(* Logix 5000 project; controller CIP vendor 1 type 14 code 106 rev 20.12; software revision 20.06; part 4 of 13 *)
(* tags used below, declared in another part *)
   Alarm_Ack : INT[8];
   Alarm_Present : INT[8];
   Alarm_Remote_Ack_All : BOOL;
   Alarm_Timer : TIMER[128];
   Bit : BOOL[128];
   IO_Status : INT;
   IO_Status_Masked : INT;
   Level_Bits : BOOL[32];
   Level_Timers : TIMER[20];
   OpCode_Pin : DINT[5];
   Recipe : RECIPE[41];
   SCLD_Dryer_Duct_Temp : REAL;
   SCLD_Solution_Tank_Lvl : REAL;
   SCLD_Supply_Flow : REAL;
   SCLD_Supply_Flow_CIP100 : REAL;
   SCLD_Supply_Flow_CIP200 : REAL;
   SCLD_Supply_Pressure : REAL;
   SCLD_Supply_Temp : REAL;
   Timer : TIMER[99];
   Timer_Chem1_Pump : TIMER[7];
   Timer_Chem2_Pump : TIMER[7];
(* MainProgram, continued *)

ROUTINE _05_ALARMS   (* ladder *)
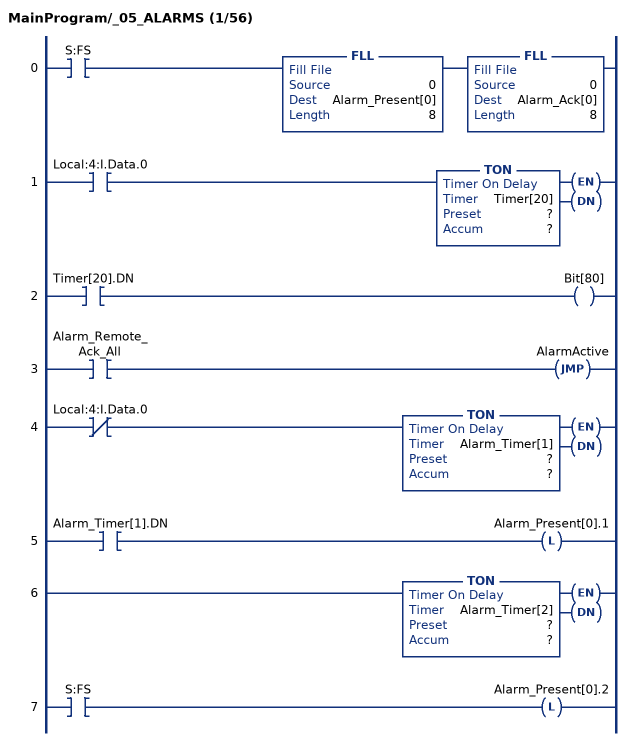
   0: XIC(S:FS)FLL(0,Alarm_Present[0],8)FLL(0,Alarm_Ack[0],8);
   1: XIC(Local:4:I.Data.0)TON(Timer[20],?,?);
   2: XIC(Timer[20].DN)OTE(Bit[80]);
   3: XIC(Alarm_Remote_Ack_All)JMP(AlarmActive);
   4: XIO(Local:4:I.Data.0)TON(Alarm_Timer[1],?,?);
   5: XIC(Alarm_Timer[1].DN)OTL(Alarm_Present[0].1);
   6: TON(Alarm_Timer[2],?,?);
   7: XIC(S:FS)OTL(Alarm_Present[0].2);
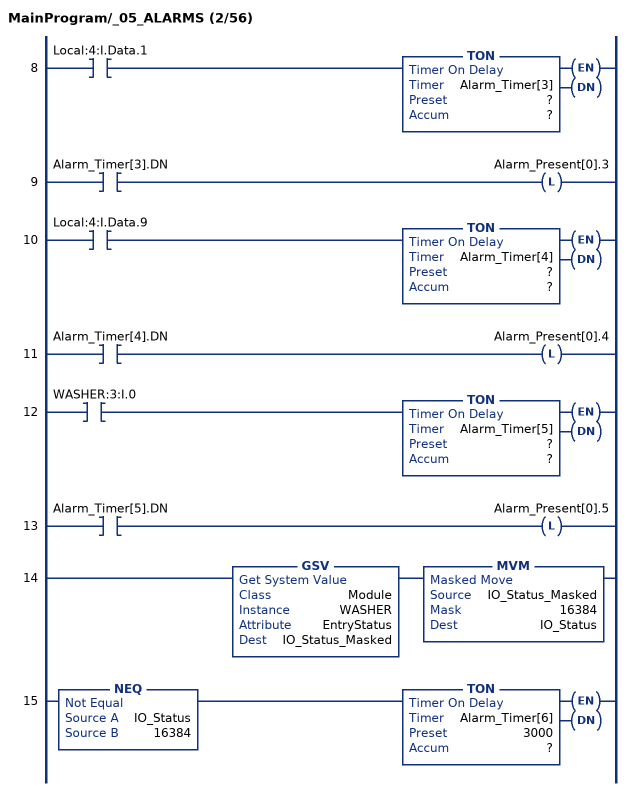
   8: XIC(Local:4:I.Data.1)TON(Alarm_Timer[3],?,?);
   9: XIC(Alarm_Timer[3].DN)OTL(Alarm_Present[0].3);
   10: XIC(Local:4:I.Data.9)TON(Alarm_Timer[4],?,?);
   11: XIC(Alarm_Timer[4].DN)OTL(Alarm_Present[0].4);
   12: XIC(WASHER:3:I.0)TON(Alarm_Timer[5],?,?);
   13: XIC(Alarm_Timer[5].DN)OTL(Alarm_Present[0].5);
   14: GSV(Module,WASHER,EntryStatus,IO_Status_Masked)MVM(IO_Status_Masked,16384,IO_Status);
   15: NEQ(IO_Status,16384)TON(Alarm_Timer[6],?,?);
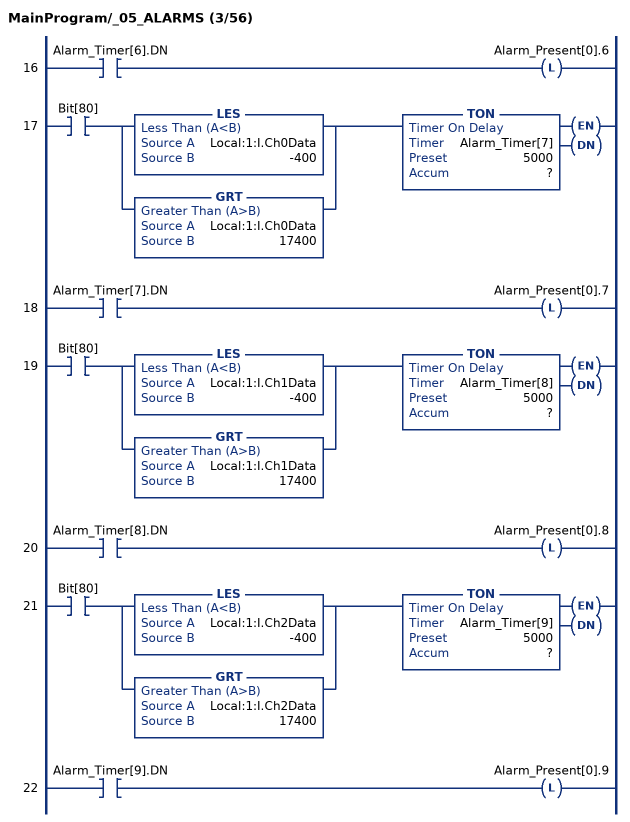
   16: XIC(Alarm_Timer[6].DN)OTL(Alarm_Present[0].6);
   17: XIC(Bit[80])[LES(Local:1:I.Ch0Data,-400) ,GRT(Local:1:I.Ch0Data,17400) ]TON(Alarm_Timer[7],?,?);
   18: XIC(Alarm_Timer[7].DN)OTL(Alarm_Present[0].7);
   19: XIC(Bit[80])[LES(Local:1:I.Ch1Data,-400) ,GRT(Local:1:I.Ch1Data,17400) ]TON(Alarm_Timer[8],?,?);
   20: XIC(Alarm_Timer[8].DN)OTL(Alarm_Present[0].8);
   21: XIC(Bit[80])[LES(Local:1:I.Ch2Data,-400) ,GRT(Local:1:I.Ch2Data,17400) ]TON(Alarm_Timer[9],?,?);
   22: XIC(Alarm_Timer[9].DN)OTL(Alarm_Present[0].9);
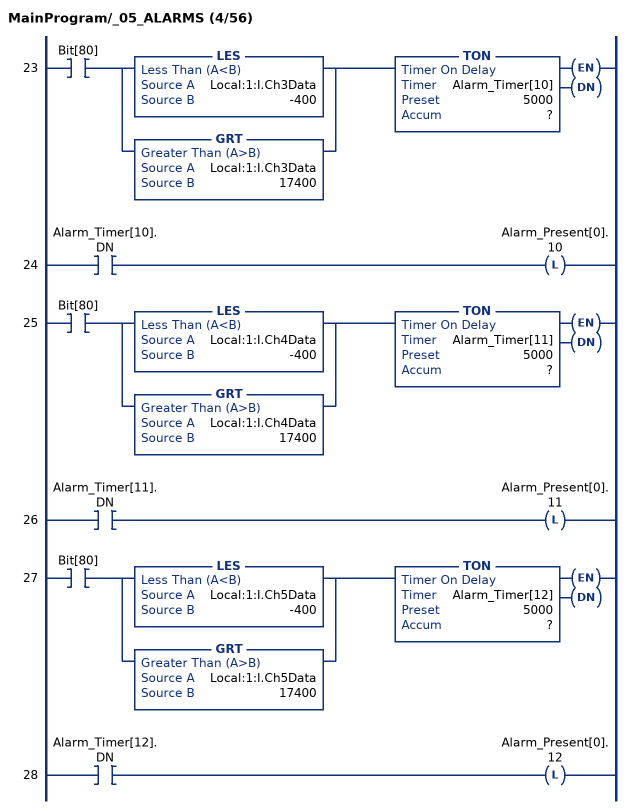
   23: XIC(Bit[80])[LES(Local:1:I.Ch3Data,-400) ,GRT(Local:1:I.Ch3Data,17400) ]TON(Alarm_Timer[10],?,?);
   24: XIC(Alarm_Timer[10].DN)OTL(Alarm_Present[0].10);
   25: XIC(Bit[80])[LES(Local:1:I.Ch4Data,-400) ,GRT(Local:1:I.Ch4Data,17400) ]TON(Alarm_Timer[11],?,?);
   26: XIC(Alarm_Timer[11].DN)OTL(Alarm_Present[0].11);
   27: XIC(Bit[80])[LES(Local:1:I.Ch5Data,-400) ,GRT(Local:1:I.Ch5Data,17400) ]TON(Alarm_Timer[12],?,?);
   28: XIC(Alarm_Timer[12].DN)OTL(Alarm_Present[0].12);
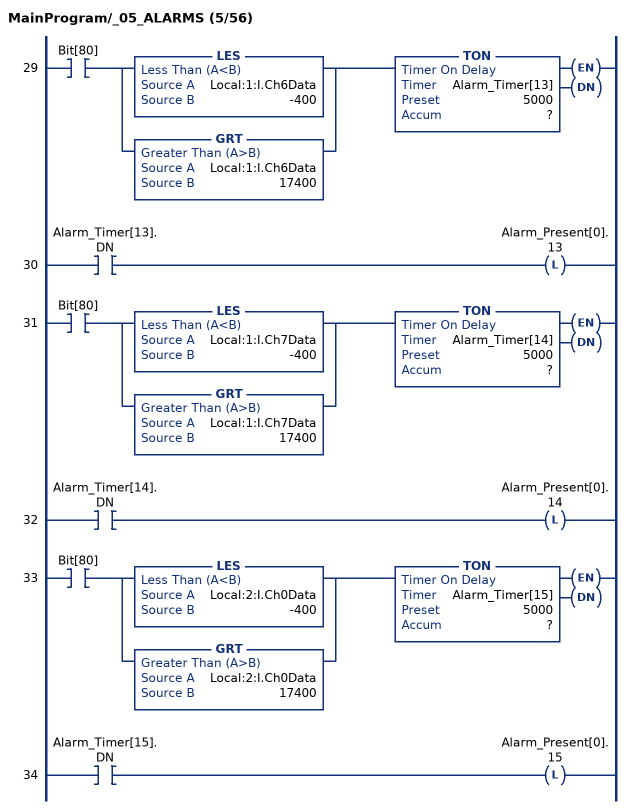
   29: XIC(Bit[80])[LES(Local:1:I.Ch6Data,-400) ,GRT(Local:1:I.Ch6Data,17400) ]TON(Alarm_Timer[13],?,?);
   30: XIC(Alarm_Timer[13].DN)OTL(Alarm_Present[0].13);
   31: XIC(Bit[80])[LES(Local:1:I.Ch7Data,-400) ,GRT(Local:1:I.Ch7Data,17400) ]TON(Alarm_Timer[14],?,?);
   32: XIC(Alarm_Timer[14].DN)OTL(Alarm_Present[0].14);
   33: XIC(Bit[80])[LES(Local:2:I.Ch0Data,-400) ,GRT(Local:2:I.Ch0Data,17400) ]TON(Alarm_Timer[15],?,?);
   34: XIC(Alarm_Timer[15].DN)OTL(Alarm_Present[0].15);
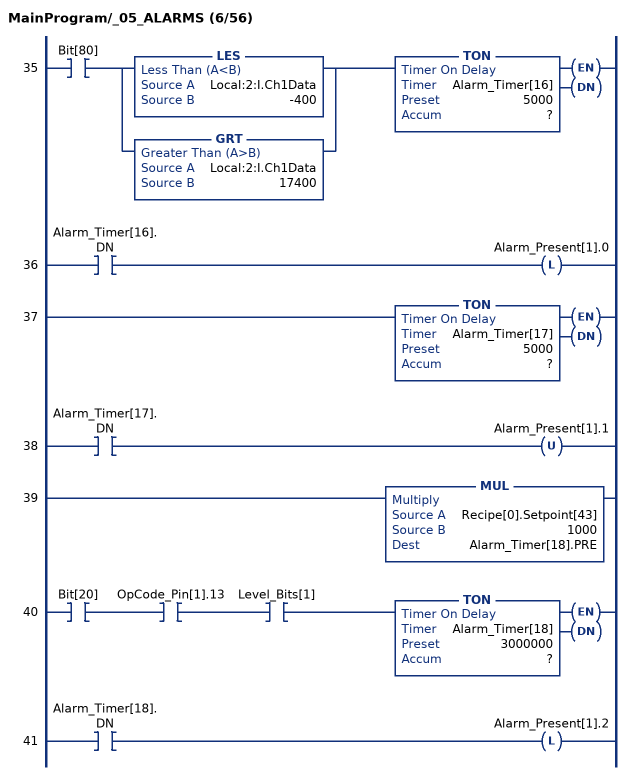
   35: XIC(Bit[80])[LES(Local:2:I.Ch1Data,-400) ,GRT(Local:2:I.Ch1Data,17400) ]TON(Alarm_Timer[16],?,?);
   36: XIC(Alarm_Timer[16].DN)OTL(Alarm_Present[1].0);
   37: TON(Alarm_Timer[17],?,?);
   38: XIC(Alarm_Timer[17].DN)OTU(Alarm_Present[1].1);
   39: MUL(Recipe[0].Setpoint[43],1000,Alarm_Timer[18].PRE);
   40: XIC(Bit[20])XIC(OpCode_Pin[1].13)XIC(Level_Bits[1])TON(Alarm_Timer[18],?,?);
   41: XIC(Alarm_Timer[18].DN)OTL(Alarm_Present[1].2);
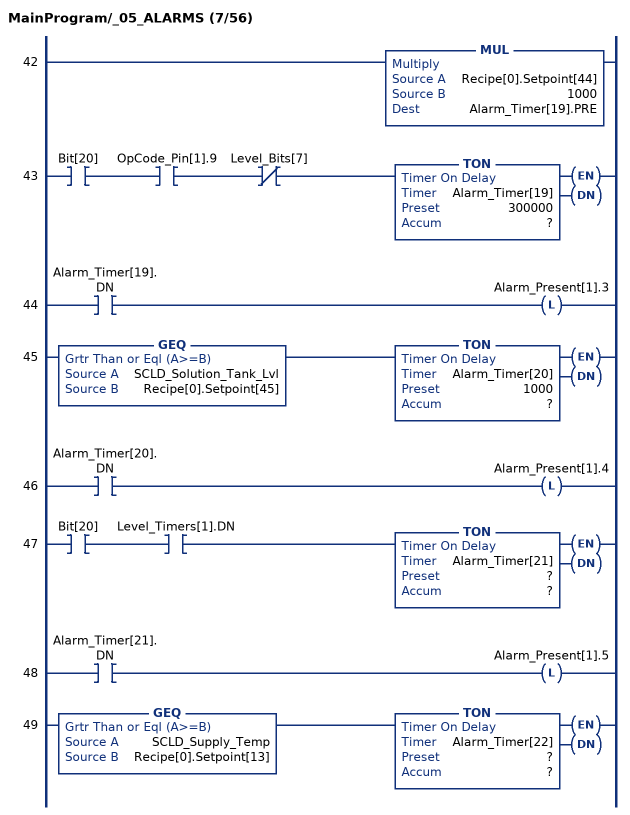
   42: MUL(Recipe[0].Setpoint[44],1000,Alarm_Timer[19].PRE);
   43: XIC(Bit[20])XIC(OpCode_Pin[1].9)XIO(Level_Bits[7])TON(Alarm_Timer[19],?,?);
   44: XIC(Alarm_Timer[19].DN)OTL(Alarm_Present[1].3);
   45: GEQ(SCLD_Solution_Tank_Lvl,Recipe[0].Setpoint[45])TON(Alarm_Timer[20],?,?);
   46: XIC(Alarm_Timer[20].DN)OTL(Alarm_Present[1].4);
   47: XIC(Bit[20])XIC(Level_Timers[1].DN)TON(Alarm_Timer[21],?,?);
   48: XIC(Alarm_Timer[21].DN)OTL(Alarm_Present[1].5);
   49: GEQ(SCLD_Supply_Temp,Recipe[0].Setpoint[13])TON(Alarm_Timer[22],?,?);
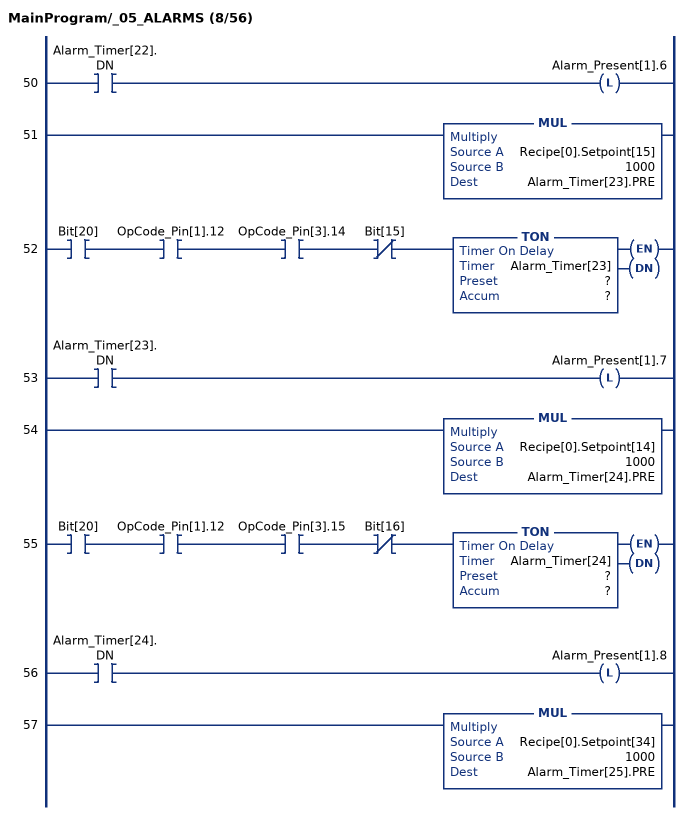
   50: XIC(Alarm_Timer[22].DN)OTL(Alarm_Present[1].6);
   51: MUL(Recipe[0].Setpoint[15],1000,Alarm_Timer[23].PRE);
   52: XIC(Bit[20])XIC(OpCode_Pin[1].12)XIC(OpCode_Pin[3].14)XIO(Bit[15])TON(Alarm_Timer[23],?,?);
   53: XIC(Alarm_Timer[23].DN)OTL(Alarm_Present[1].7);
   54: MUL(Recipe[0].Setpoint[14],1000,Alarm_Timer[24].PRE);
   55: XIC(Bit[20])XIC(OpCode_Pin[1].12)XIC(OpCode_Pin[3].15)XIO(Bit[16])TON(Alarm_Timer[24],?,?);
   56: XIC(Alarm_Timer[24].DN)OTL(Alarm_Present[1].8);
   57: MUL(Recipe[0].Setpoint[34],1000,Alarm_Timer[25].PRE);
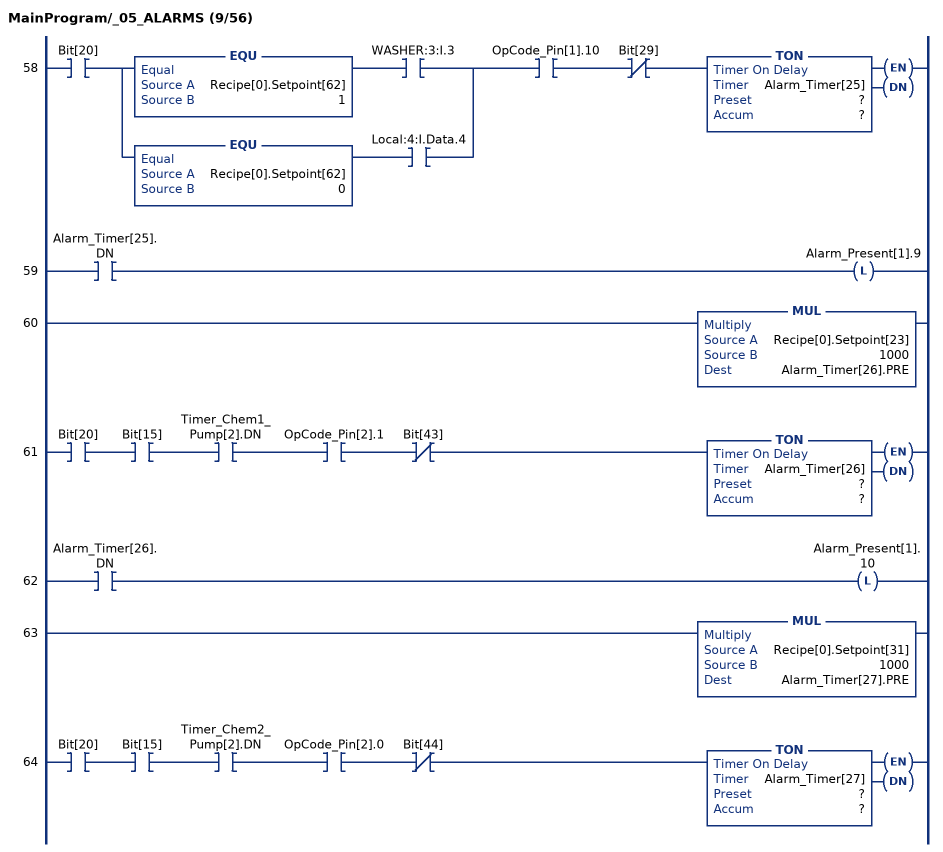
   58: XIC(Bit[20])[EQU(Recipe[0].Setpoint[62],1) XIC(WASHER:3:I.3) ,EQU(Recipe[0].Setpoint[62],0) XIC(Local:4:I.Data.4) ]XIC(OpCode_Pin[1].10)XIO(Bit[29])TON(Alarm_Timer[25],?,?);
   59: XIC(Alarm_Timer[25].DN)OTL(Alarm_Present[1].9);
   60: MUL(Recipe[0].Setpoint[23],1000,Alarm_Timer[26].PRE);
   61: XIC(Bit[20])XIC(Bit[15])XIC(Timer_Chem1_Pump[2].DN)XIC(OpCode_Pin[2].1)XIO(Bit[43])TON(Alarm_Timer[26],?,?);
   62: XIC(Alarm_Timer[26].DN)OTL(Alarm_Present[1].10);
   63: MUL(Recipe[0].Setpoint[31],1000,Alarm_Timer[27].PRE);
   64: XIC(Bit[20])XIC(Bit[15])XIC(Timer_Chem2_Pump[2].DN)XIC(OpCode_Pin[2].0)XIO(Bit[44])TON(Alarm_Timer[27],?,?);
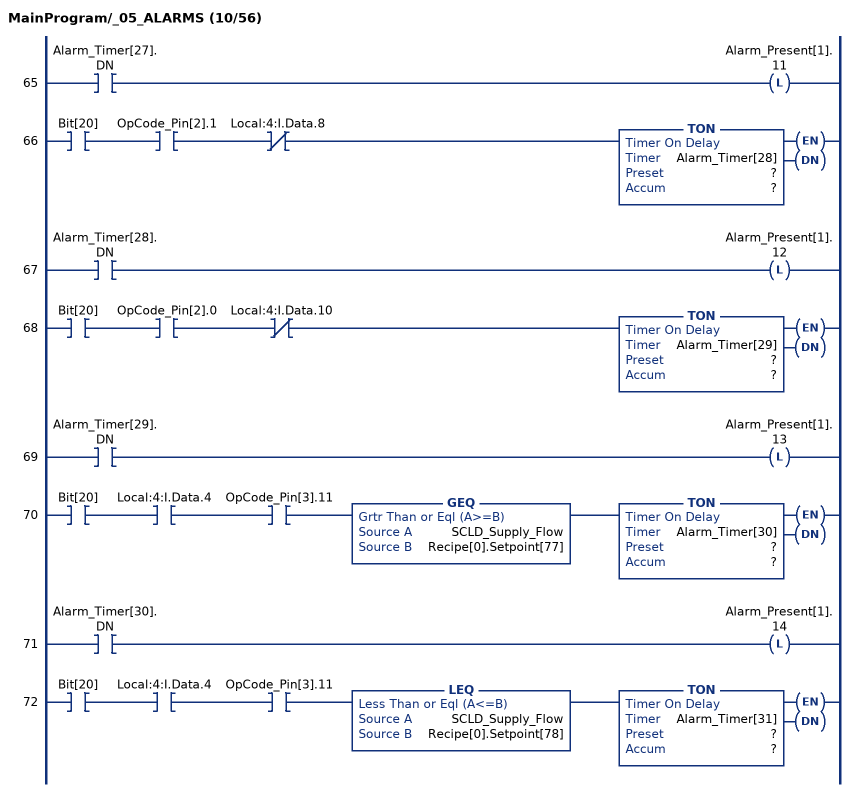
   65: XIC(Alarm_Timer[27].DN)OTL(Alarm_Present[1].11);
   66: XIC(Bit[20])XIC(OpCode_Pin[2].1)XIO(Local:4:I.Data.8)TON(Alarm_Timer[28],?,?);
   67: XIC(Alarm_Timer[28].DN)OTL(Alarm_Present[1].12);
   68: XIC(Bit[20])XIC(OpCode_Pin[2].0)XIO(Local:4:I.Data.10)TON(Alarm_Timer[29],?,?);
   69: XIC(Alarm_Timer[29].DN)OTL(Alarm_Present[1].13);
   70: XIC(Bit[20])XIC(Local:4:I.Data.4)XIC(OpCode_Pin[3].11)GEQ(SCLD_Supply_Flow,Recipe[0].Setpoint[77])TON(Alarm_Timer[30],?,?);
   71: XIC(Alarm_Timer[30].DN)OTL(Alarm_Present[1].14);
   72: XIC(Bit[20])XIC(Local:4:I.Data.4)XIC(OpCode_Pin[3].11)LEQ(SCLD_Supply_Flow,Recipe[0].Setpoint[78])TON(Alarm_Timer[31],?,?);
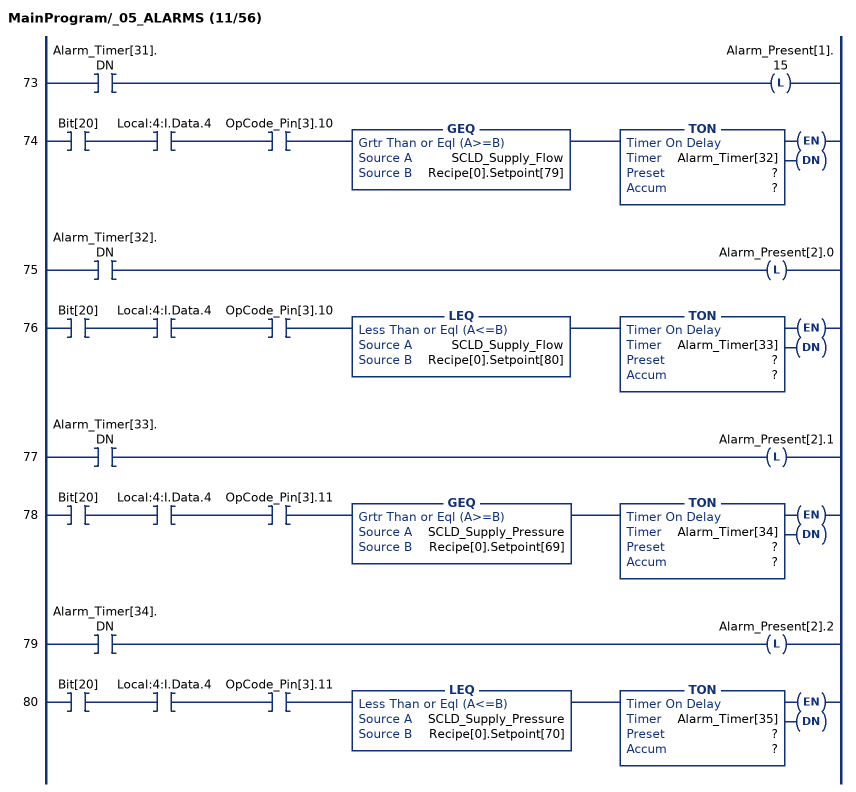
   73: XIC(Alarm_Timer[31].DN)OTL(Alarm_Present[1].15);
   74: XIC(Bit[20])XIC(Local:4:I.Data.4)XIC(OpCode_Pin[3].10)GEQ(SCLD_Supply_Flow,Recipe[0].Setpoint[79])TON(Alarm_Timer[32],?,?);
   75: XIC(Alarm_Timer[32].DN)OTL(Alarm_Present[2].0);
   76: XIC(Bit[20])XIC(Local:4:I.Data.4)XIC(OpCode_Pin[3].10)LEQ(SCLD_Supply_Flow,Recipe[0].Setpoint[80])TON(Alarm_Timer[33],?,?);
   77: XIC(Alarm_Timer[33].DN)OTL(Alarm_Present[2].1);
   78: XIC(Bit[20])XIC(Local:4:I.Data.4)XIC(OpCode_Pin[3].11)GEQ(SCLD_Supply_Pressure,Recipe[0].Setpoint[69])TON(Alarm_Timer[34],?,?);
   79: XIC(Alarm_Timer[34].DN)OTL(Alarm_Present[2].2);
   80: XIC(Bit[20])XIC(Local:4:I.Data.4)XIC(OpCode_Pin[3].11)LEQ(SCLD_Supply_Pressure,Recipe[0].Setpoint[70])TON(Alarm_Timer[35],?,?);
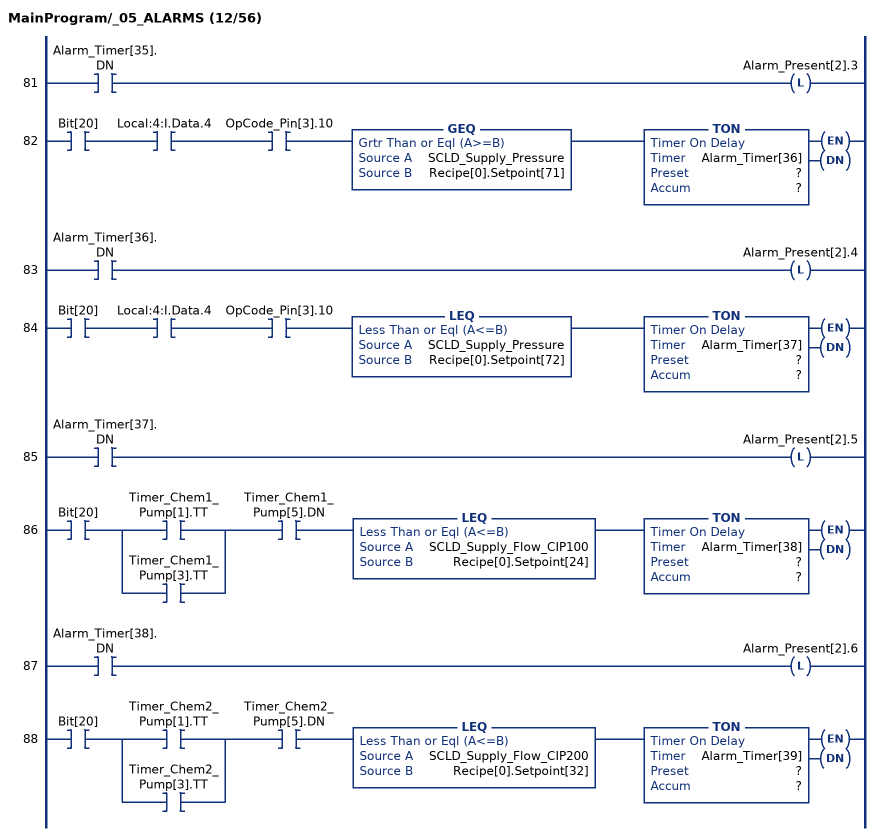
   81: XIC(Alarm_Timer[35].DN)OTL(Alarm_Present[2].3);
   82: XIC(Bit[20])XIC(Local:4:I.Data.4)XIC(OpCode_Pin[3].10)GEQ(SCLD_Supply_Pressure,Recipe[0].Setpoint[71])TON(Alarm_Timer[36],?,?);
   83: XIC(Alarm_Timer[36].DN)OTL(Alarm_Present[2].4);
   84: XIC(Bit[20])XIC(Local:4:I.Data.4)XIC(OpCode_Pin[3].10)LEQ(SCLD_Supply_Pressure,Recipe[0].Setpoint[72])TON(Alarm_Timer[37],?,?);
   85: XIC(Alarm_Timer[37].DN)OTL(Alarm_Present[2].5);
   86: XIC(Bit[20])[XIC(Timer_Chem1_Pump[1].TT) ,XIC(Timer_Chem1_Pump[3].TT) ]XIC(Timer_Chem1_Pump[5].DN)LEQ(SCLD_Supply_Flow_CIP100,Recipe[0].Setpoint[24])TON(Alarm_Timer[38],?,?);
   87: XIC(Alarm_Timer[38].DN)OTL(Alarm_Present[2].6);
   88: XIC(Bit[20])[XIC(Timer_Chem2_Pump[1].TT) ,XIC(Timer_Chem2_Pump[3].TT) ]XIC(Timer_Chem2_Pump[5].DN)LEQ(SCLD_Supply_Flow_CIP200,Recipe[0].Setpoint[32])TON(Alarm_Timer[39],?,?);
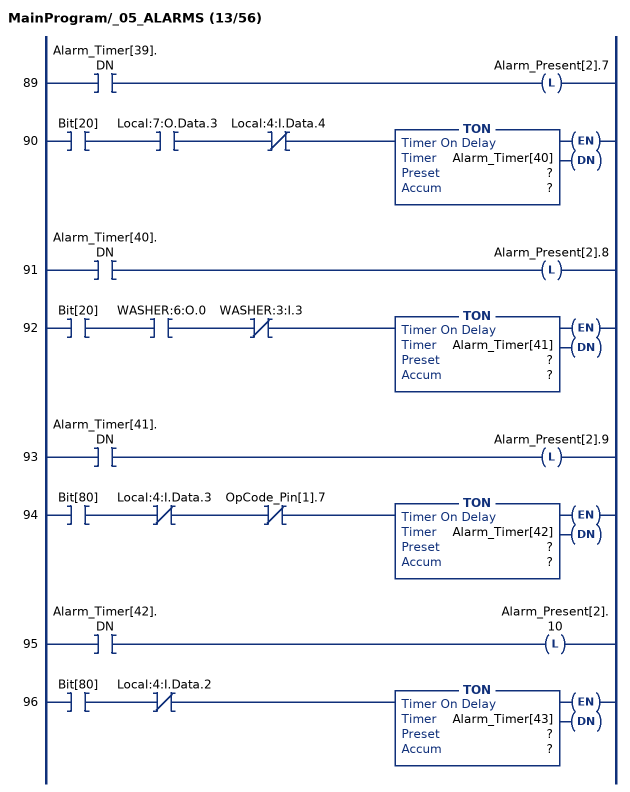
   89: XIC(Alarm_Timer[39].DN)OTL(Alarm_Present[2].7);
   90: XIC(Bit[20])XIC(Local:7:O.Data.3)XIO(Local:4:I.Data.4)TON(Alarm_Timer[40],?,?);
   91: XIC(Alarm_Timer[40].DN)OTL(Alarm_Present[2].8);
   92: XIC(Bit[20])XIC(WASHER:6:O.0)XIO(WASHER:3:I.3)TON(Alarm_Timer[41],?,?);
   93: XIC(Alarm_Timer[41].DN)OTL(Alarm_Present[2].9);
   94: XIC(Bit[80])XIO(Local:4:I.Data.3)XIO(OpCode_Pin[1].7)TON(Alarm_Timer[42],?,?);
   95: XIC(Alarm_Timer[42].DN)OTL(Alarm_Present[2].10);
   96: XIC(Bit[80])XIO(Local:4:I.Data.2)TON(Alarm_Timer[43],?,?);
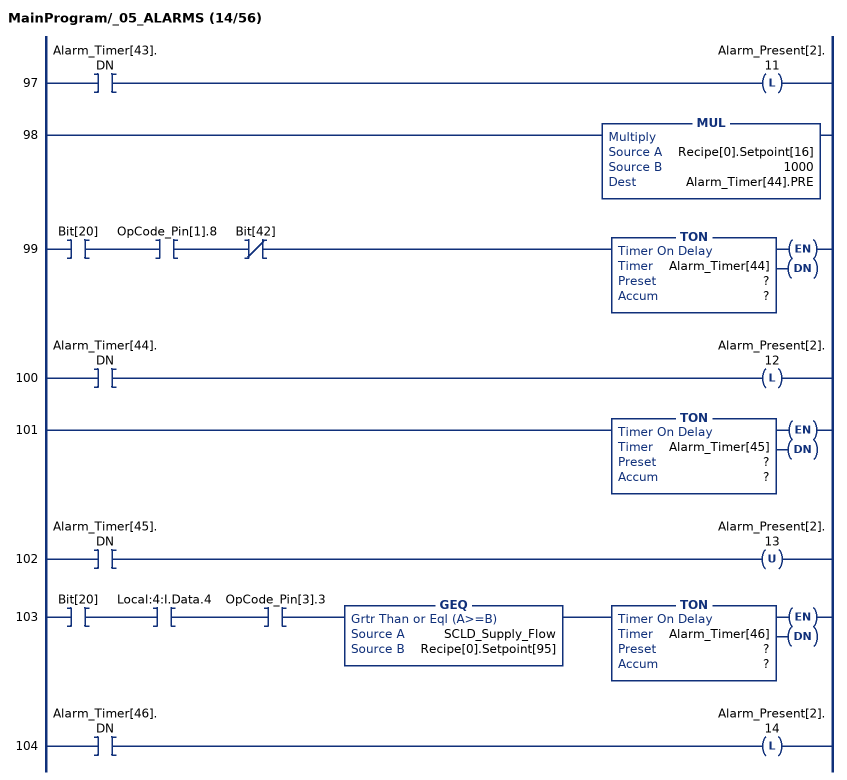
   97: XIC(Alarm_Timer[43].DN)OTL(Alarm_Present[2].11);
   98: MUL(Recipe[0].Setpoint[16],1000,Alarm_Timer[44].PRE);
   99: XIC(Bit[20])XIC(OpCode_Pin[1].8)XIO(Bit[42])TON(Alarm_Timer[44],?,?);
   100: XIC(Alarm_Timer[44].DN)OTL(Alarm_Present[2].12);
   101: TON(Alarm_Timer[45],?,?);
   102: XIC(Alarm_Timer[45].DN)OTU(Alarm_Present[2].13);
   103: XIC(Bit[20])XIC(Local:4:I.Data.4)XIC(OpCode_Pin[3].3)GEQ(SCLD_Supply_Flow,Recipe[0].Setpoint[95])TON(Alarm_Timer[46],?,?);
   104: XIC(Alarm_Timer[46].DN)OTL(Alarm_Present[2].14);
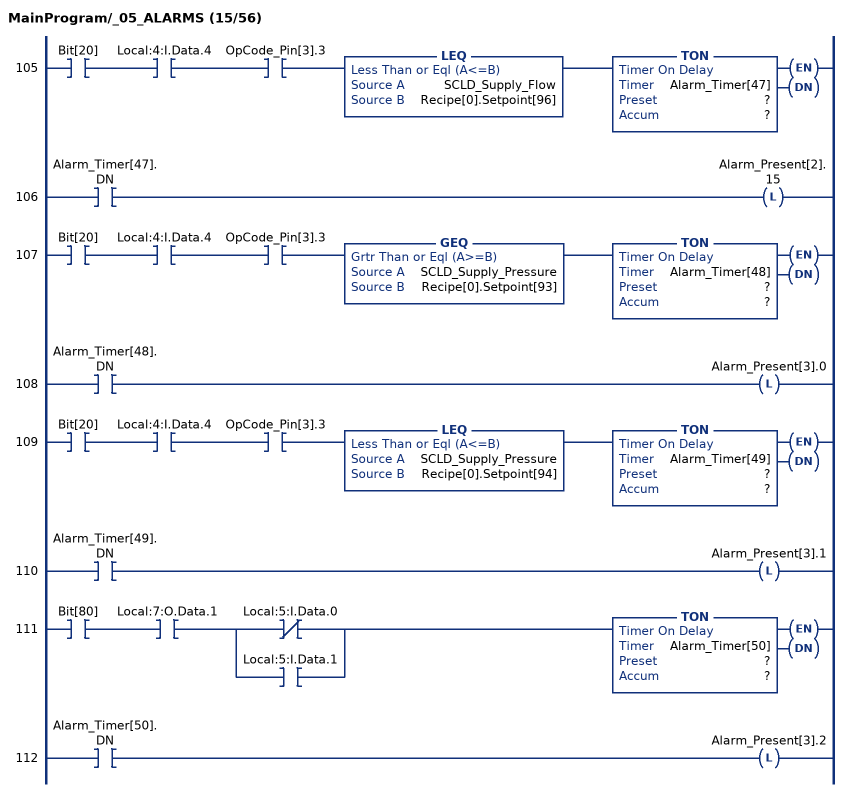
   105: XIC(Bit[20])XIC(Local:4:I.Data.4)XIC(OpCode_Pin[3].3)LEQ(SCLD_Supply_Flow,Recipe[0].Setpoint[96])TON(Alarm_Timer[47],?,?);
   106: XIC(Alarm_Timer[47].DN)OTL(Alarm_Present[2].15);
   107: XIC(Bit[20])XIC(Local:4:I.Data.4)XIC(OpCode_Pin[3].3)GEQ(SCLD_Supply_Pressure,Recipe[0].Setpoint[93])TON(Alarm_Timer[48],?,?);
   108: XIC(Alarm_Timer[48].DN)OTL(Alarm_Present[3].0);
   109: XIC(Bit[20])XIC(Local:4:I.Data.4)XIC(OpCode_Pin[3].3)LEQ(SCLD_Supply_Pressure,Recipe[0].Setpoint[94])TON(Alarm_Timer[49],?,?);
   110: XIC(Alarm_Timer[49].DN)OTL(Alarm_Present[3].1);
   111: XIC(Bit[80])XIC(Local:7:O.Data.1)[XIO(Local:5:I.Data.0) ,XIC(Local:5:I.Data.1) ]TON(Alarm_Timer[50],?,?);
   112: XIC(Alarm_Timer[50].DN)OTL(Alarm_Present[3].2);
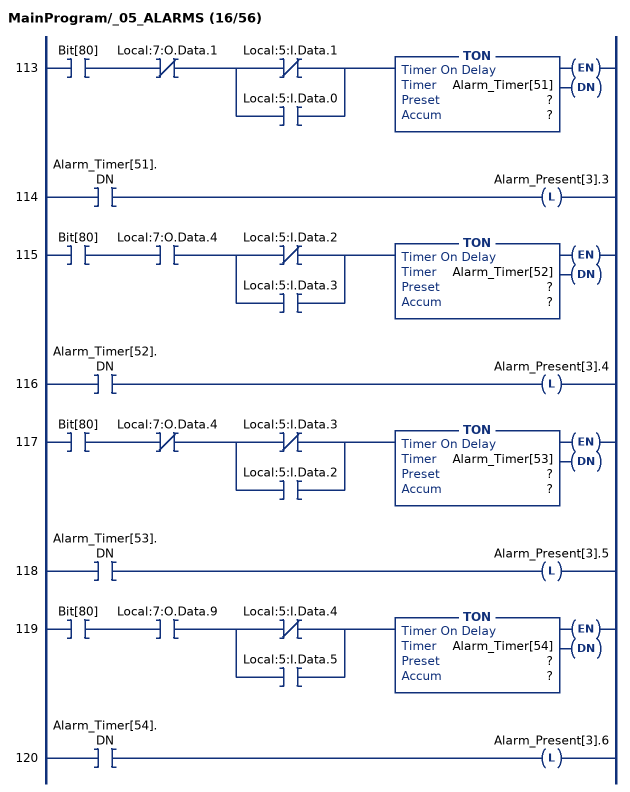
   113: XIC(Bit[80])XIO(Local:7:O.Data.1)[XIO(Local:5:I.Data.1) ,XIC(Local:5:I.Data.0) ]TON(Alarm_Timer[51],?,?);
   114: XIC(Alarm_Timer[51].DN)OTL(Alarm_Present[3].3);
   115: XIC(Bit[80])XIC(Local:7:O.Data.4)[XIO(Local:5:I.Data.2) ,XIC(Local:5:I.Data.3) ]TON(Alarm_Timer[52],?,?);
   116: XIC(Alarm_Timer[52].DN)OTL(Alarm_Present[3].4);
   117: XIC(Bit[80])XIO(Local:7:O.Data.4)[XIO(Local:5:I.Data.3) ,XIC(Local:5:I.Data.2) ]TON(Alarm_Timer[53],?,?);
   118: XIC(Alarm_Timer[53].DN)OTL(Alarm_Present[3].5);
   119: XIC(Bit[80])XIC(Local:7:O.Data.9)[XIO(Local:5:I.Data.4) ,XIC(Local:5:I.Data.5) ]TON(Alarm_Timer[54],?,?);
   120: XIC(Alarm_Timer[54].DN)OTL(Alarm_Present[3].6);
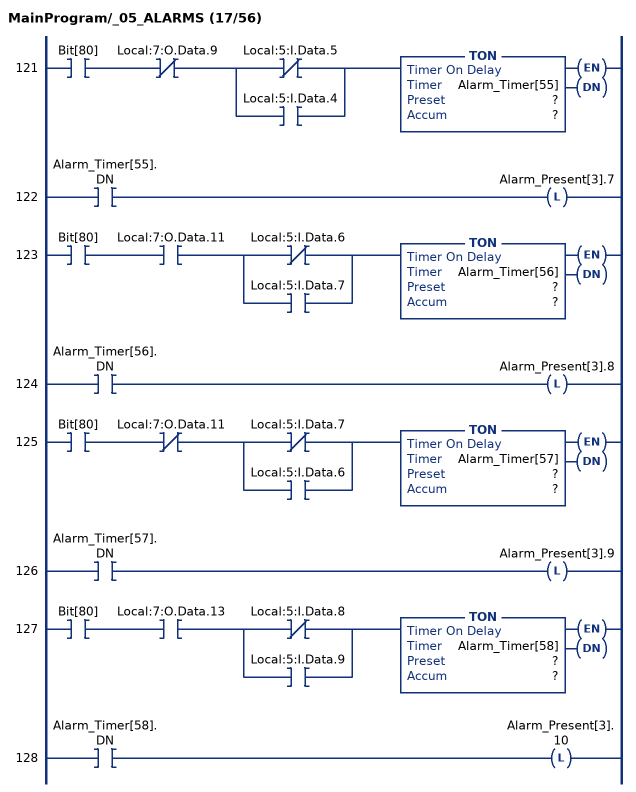
   121: XIC(Bit[80])XIO(Local:7:O.Data.9)[XIO(Local:5:I.Data.5) ,XIC(Local:5:I.Data.4) ]TON(Alarm_Timer[55],?,?);
   122: XIC(Alarm_Timer[55].DN)OTL(Alarm_Present[3].7);
   123: XIC(Bit[80])XIC(Local:7:O.Data.11)[XIO(Local:5:I.Data.6) ,XIC(Local:5:I.Data.7) ]TON(Alarm_Timer[56],?,?);
   124: XIC(Alarm_Timer[56].DN)OTL(Alarm_Present[3].8);
   125: XIC(Bit[80])XIO(Local:7:O.Data.11)[XIO(Local:5:I.Data.7) ,XIC(Local:5:I.Data.6) ]TON(Alarm_Timer[57],?,?);
   126: XIC(Alarm_Timer[57].DN)OTL(Alarm_Present[3].9);
   127: XIC(Bit[80])XIC(Local:7:O.Data.13)[XIO(Local:5:I.Data.8) ,XIC(Local:5:I.Data.9) ]TON(Alarm_Timer[58],?,?);
   128: XIC(Alarm_Timer[58].DN)OTL(Alarm_Present[3].10);
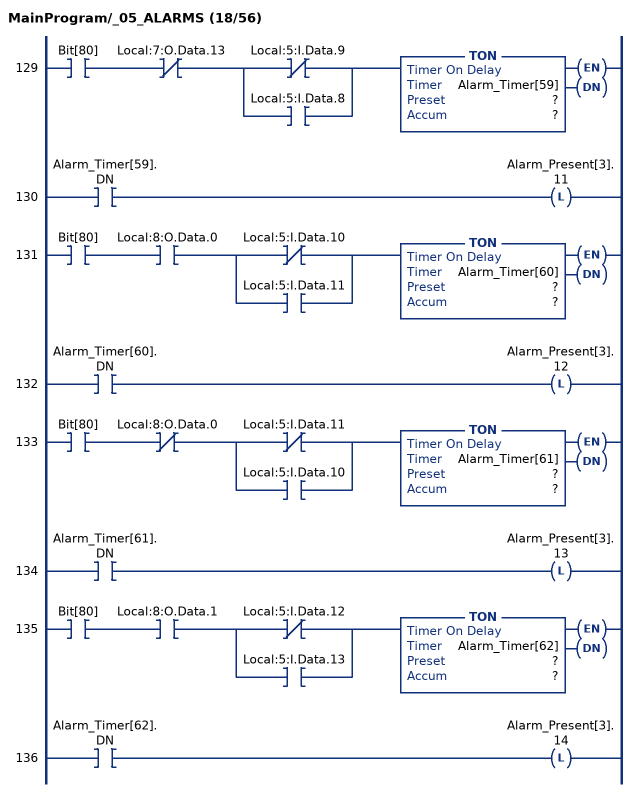
   129: XIC(Bit[80])XIO(Local:7:O.Data.13)[XIO(Local:5:I.Data.9) ,XIC(Local:5:I.Data.8) ]TON(Alarm_Timer[59],?,?);
   130: XIC(Alarm_Timer[59].DN)OTL(Alarm_Present[3].11);
   131: XIC(Bit[80])XIC(Local:8:O.Data.0)[XIO(Local:5:I.Data.10) ,XIC(Local:5:I.Data.11) ]TON(Alarm_Timer[60],?,?);
   132: XIC(Alarm_Timer[60].DN)OTL(Alarm_Present[3].12);
   133: XIC(Bit[80])XIO(Local:8:O.Data.0)[XIO(Local:5:I.Data.11) ,XIC(Local:5:I.Data.10) ]TON(Alarm_Timer[61],?,?);
   134: XIC(Alarm_Timer[61].DN)OTL(Alarm_Present[3].13);
   135: XIC(Bit[80])XIC(Local:8:O.Data.1)[XIO(Local:5:I.Data.12) ,XIC(Local:5:I.Data.13) ]TON(Alarm_Timer[62],?,?);
   136: XIC(Alarm_Timer[62].DN)OTL(Alarm_Present[3].14);
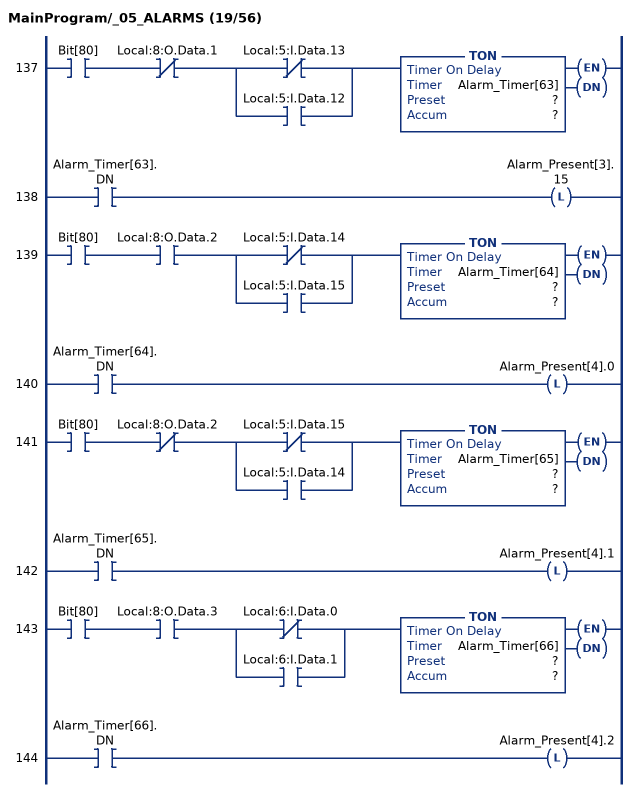
   137: XIC(Bit[80])XIO(Local:8:O.Data.1)[XIO(Local:5:I.Data.13) ,XIC(Local:5:I.Data.12) ]TON(Alarm_Timer[63],?,?);
   138: XIC(Alarm_Timer[63].DN)OTL(Alarm_Present[3].15);
   139: XIC(Bit[80])XIC(Local:8:O.Data.2)[XIO(Local:5:I.Data.14) ,XIC(Local:5:I.Data.15) ]TON(Alarm_Timer[64],?,?);
   140: XIC(Alarm_Timer[64].DN)OTL(Alarm_Present[4].0);
   141: XIC(Bit[80])XIO(Local:8:O.Data.2)[XIO(Local:5:I.Data.15) ,XIC(Local:5:I.Data.14) ]TON(Alarm_Timer[65],?,?);
   142: XIC(Alarm_Timer[65].DN)OTL(Alarm_Present[4].1);
   143: XIC(Bit[80])XIC(Local:8:O.Data.3)[XIO(Local:6:I.Data.0) ,XIC(Local:6:I.Data.1) ]TON(Alarm_Timer[66],?,?);
   144: XIC(Alarm_Timer[66].DN)OTL(Alarm_Present[4].2);
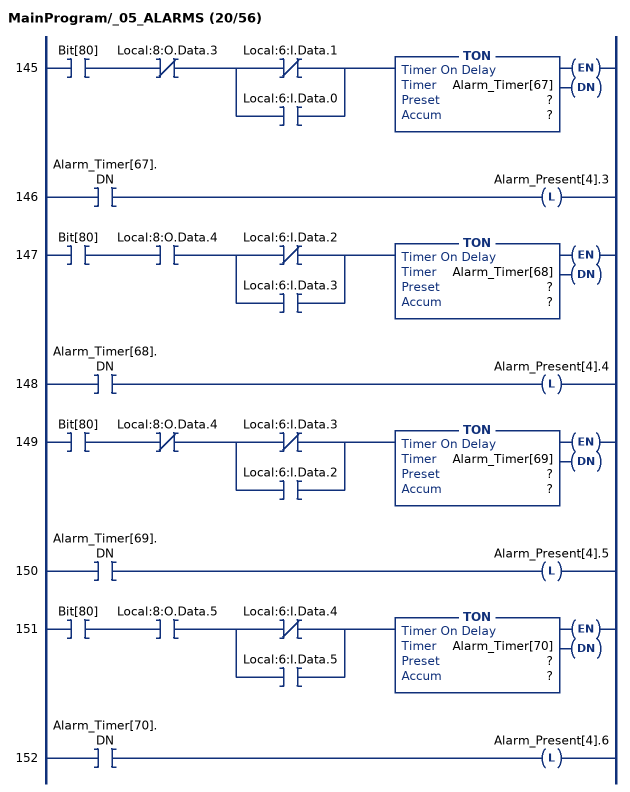
   145: XIC(Bit[80])XIO(Local:8:O.Data.3)[XIO(Local:6:I.Data.1) ,XIC(Local:6:I.Data.0) ]TON(Alarm_Timer[67],?,?);
   146: XIC(Alarm_Timer[67].DN)OTL(Alarm_Present[4].3);
   147: XIC(Bit[80])XIC(Local:8:O.Data.4)[XIO(Local:6:I.Data.2) ,XIC(Local:6:I.Data.3) ]TON(Alarm_Timer[68],?,?);
   148: XIC(Alarm_Timer[68].DN)OTL(Alarm_Present[4].4);
   149: XIC(Bit[80])XIO(Local:8:O.Data.4)[XIO(Local:6:I.Data.3) ,XIC(Local:6:I.Data.2) ]TON(Alarm_Timer[69],?,?);
   150: XIC(Alarm_Timer[69].DN)OTL(Alarm_Present[4].5);
   151: XIC(Bit[80])XIC(Local:8:O.Data.5)[XIO(Local:6:I.Data.4) ,XIC(Local:6:I.Data.5) ]TON(Alarm_Timer[70],?,?);
   152: XIC(Alarm_Timer[70].DN)OTL(Alarm_Present[4].6);
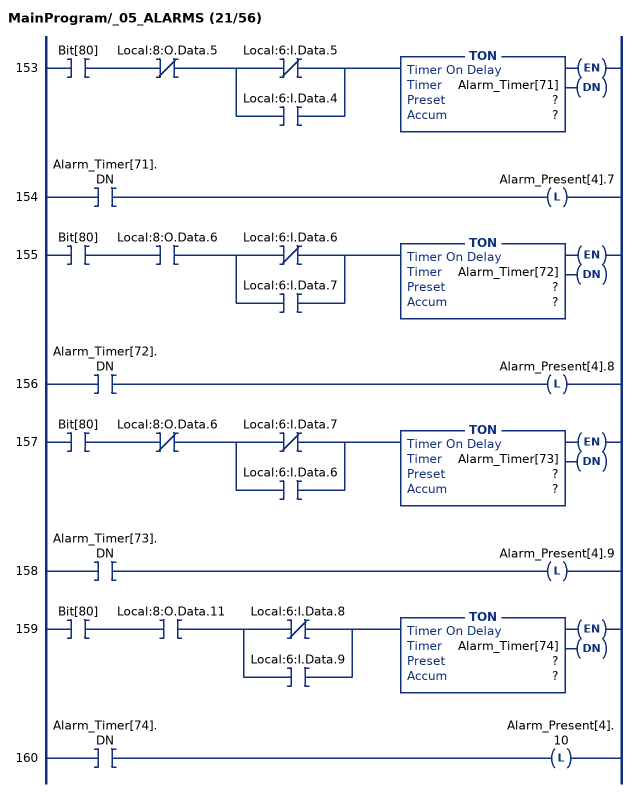
   153: XIC(Bit[80])XIO(Local:8:O.Data.5)[XIO(Local:6:I.Data.5) ,XIC(Local:6:I.Data.4) ]TON(Alarm_Timer[71],?,?);
   154: XIC(Alarm_Timer[71].DN)OTL(Alarm_Present[4].7);
   155: XIC(Bit[80])XIC(Local:8:O.Data.6)[XIO(Local:6:I.Data.6) ,XIC(Local:6:I.Data.7) ]TON(Alarm_Timer[72],?,?);
   156: XIC(Alarm_Timer[72].DN)OTL(Alarm_Present[4].8);
   157: XIC(Bit[80])XIO(Local:8:O.Data.6)[XIO(Local:6:I.Data.7) ,XIC(Local:6:I.Data.6) ]TON(Alarm_Timer[73],?,?);
   158: XIC(Alarm_Timer[73].DN)OTL(Alarm_Present[4].9);
   159: XIC(Bit[80])XIC(Local:8:O.Data.11)[XIO(Local:6:I.Data.8) ,XIC(Local:6:I.Data.9) ]TON(Alarm_Timer[74],?,?);
   160: XIC(Alarm_Timer[74].DN)OTL(Alarm_Present[4].10);
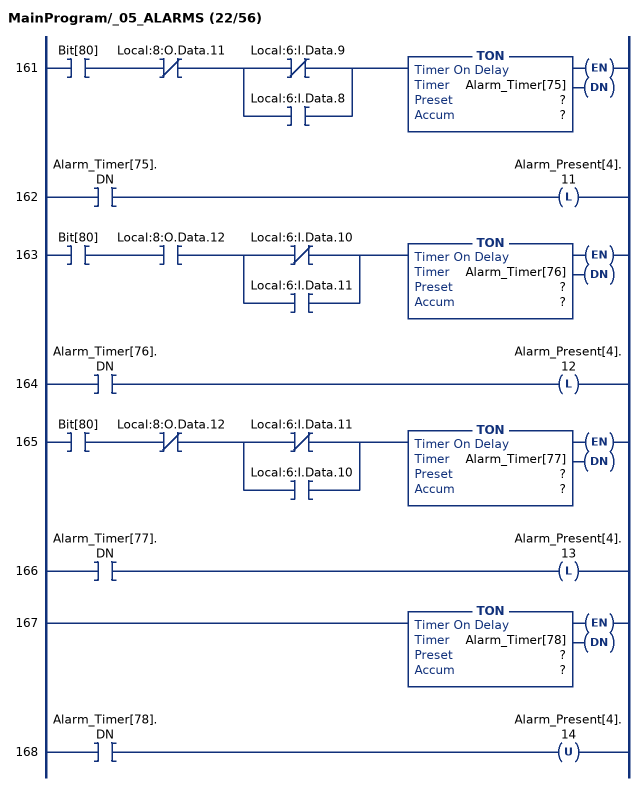
   161: XIC(Bit[80])XIO(Local:8:O.Data.11)[XIO(Local:6:I.Data.9) ,XIC(Local:6:I.Data.8) ]TON(Alarm_Timer[75],?,?);
   162: XIC(Alarm_Timer[75].DN)OTL(Alarm_Present[4].11);
   163: XIC(Bit[80])XIC(Local:8:O.Data.12)[XIO(Local:6:I.Data.10) ,XIC(Local:6:I.Data.11) ]TON(Alarm_Timer[76],?,?);
   164: XIC(Alarm_Timer[76].DN)OTL(Alarm_Present[4].12);
   165: XIC(Bit[80])XIO(Local:8:O.Data.12)[XIO(Local:6:I.Data.11) ,XIC(Local:6:I.Data.10) ]TON(Alarm_Timer[77],?,?);
   166: XIC(Alarm_Timer[77].DN)OTL(Alarm_Present[4].13);
   167: TON(Alarm_Timer[78],?,?);
   168: XIC(Alarm_Timer[78].DN)OTU(Alarm_Present[4].14);
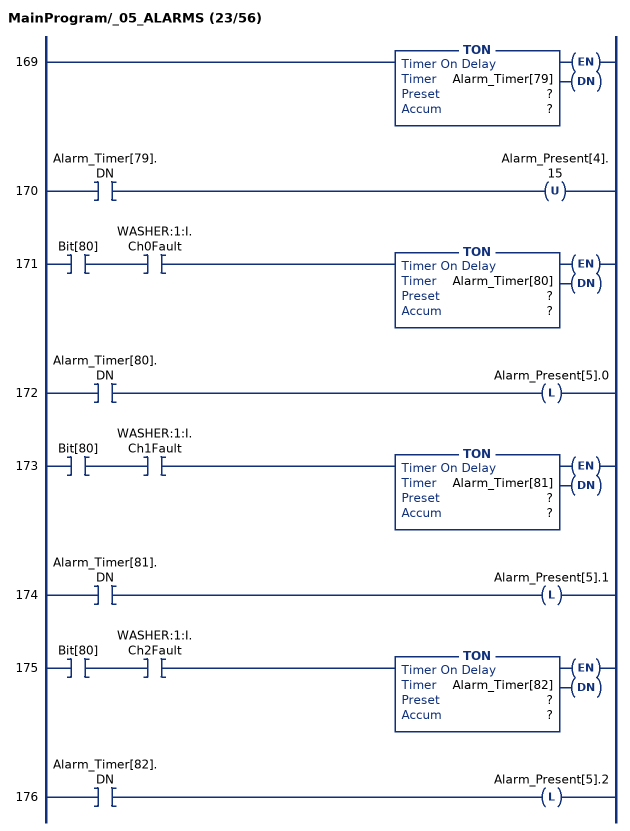
   169: TON(Alarm_Timer[79],?,?);
   170: XIC(Alarm_Timer[79].DN)OTU(Alarm_Present[4].15);
   171: XIC(Bit[80])XIC(WASHER:1:I.Ch0Fault)TON(Alarm_Timer[80],?,?);
   172: XIC(Alarm_Timer[80].DN)OTL(Alarm_Present[5].0);
   173: XIC(Bit[80])XIC(WASHER:1:I.Ch1Fault)TON(Alarm_Timer[81],?,?);
   174: XIC(Alarm_Timer[81].DN)OTL(Alarm_Present[5].1);
   175: XIC(Bit[80])XIC(WASHER:1:I.Ch2Fault)TON(Alarm_Timer[82],?,?);
   176: XIC(Alarm_Timer[82].DN)OTL(Alarm_Present[5].2);
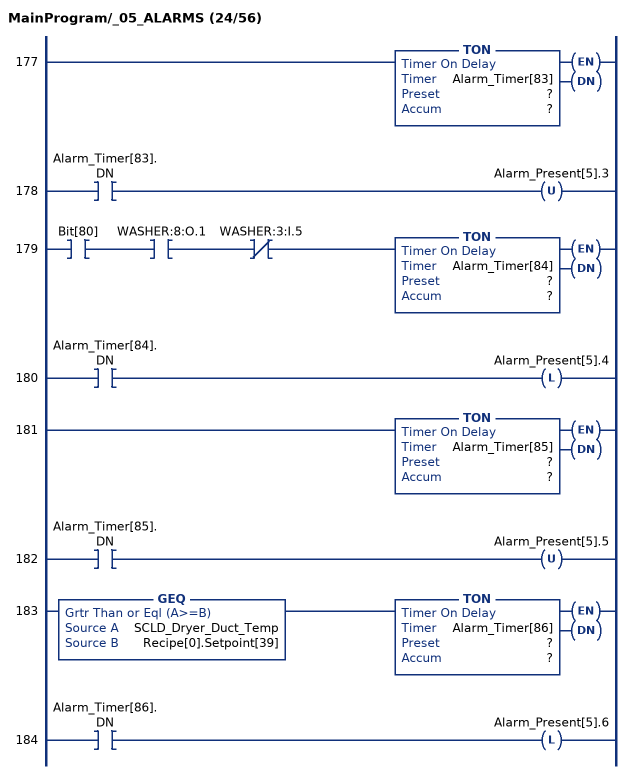
   177: TON(Alarm_Timer[83],?,?);
   178: XIC(Alarm_Timer[83].DN)OTU(Alarm_Present[5].3);
   179: XIC(Bit[80])XIC(WASHER:8:O.1)XIO(WASHER:3:I.5)TON(Alarm_Timer[84],?,?);
   180: XIC(Alarm_Timer[84].DN)OTL(Alarm_Present[5].4);
   181: TON(Alarm_Timer[85],?,?);
   182: XIC(Alarm_Timer[85].DN)OTU(Alarm_Present[5].5);
   183: GEQ(SCLD_Dryer_Duct_Temp,Recipe[0].Setpoint[39])TON(Alarm_Timer[86],?,?);
   184: XIC(Alarm_Timer[86].DN)OTL(Alarm_Present[5].6);
